Fanuc KAREL source: kt00065.KL

-- PROVISIONAL review KL for V770-1; original PC SHA256 1d701109c9aed1bf9f79d834c400fce812b98e8d73a46e65118f4a1c2bc11f15
-- Incomplete behavior may be omitted. Consult companion uncertainty JSON. Do not deploy.
PROGRAM KT00065
%NOLOCKGROUP
VAR
  I1 : INTEGER
  I2 : INTEGER
  OUT : INTEGER
BEGIN
  -- UNRESOLVED_PC offsets 5-16; opcodes 2E,23
  -- UNRESOLVED_PC offsets 21-32; opcodes 2E,23
  -- UNRESOLVED_PC offsets 37-48; opcodes 2E,23
  -- UNRESOLVED_PC offsets 53-64; opcodes 2E,23
  -- UNRESOLVED_PC offsets 69-88; opcodes 21,21,54,23
  -- UNRESOLVED_PC offsets 93-97; opcodes 7F
END KT00065
